(* PLC project station_cds.project, CODESYS CODESYS V3.5 SP22 Patch 1 *)
(* stored: creationDateTime 2026-11-25T17:27:32.1859428, modificationDateTime 2026-11-25T17:27:31.3827148 *)

FUNCTION_BLOCK FB_CurveEval
  VAR_INPUT
    Reset : BOOL;  (* clear all results, before a new pull *)
    Sample : BOOL;  (* X and F are a new sample *)
    Stroke : INT;  (* 1 pull, 2 return *)
    X : REAL;  (* mm, travel from touch *)
    F : REAL;  (* N *)
    Finish : BOOL;  (* return stroke finished: judge *)
    Mode : INT := 3;
    GateX : REAL := 3.0;  (* mm *)
    Gate2X : REAL := 10.0;  (* mm *)
    PeakXLo : REAL := 13.0;  (* mm *)
    PeakXHi : REAL := 26.0;  (* mm *)
    StepSpan : REAL := 2.0;  (* mm *)
    StopF : REAL := 30.0;  (* N *)
    G1Lo : REAL;  (* N, limits of FpG1 (mode 2) *)
    G1Hi : REAL;
    MeanLo : REAL;  (* N, limits of FMean (mode 3) *)
    MeanHi : REAL;
    HystLo : REAL;  (* N, limits of FHyst (mode 3) *)
    HystHi : REAL;
    RetFMin : REAL;  (* N, FrG1 must be above (mode 3) *)
    G2Lo : REAL;  (* N, limits of FpG2 *)
    G2Hi : REAL;
    PeakFLo : REAL;  (* N *)
    PeakFHi : REAL;
    PeakXMin : REAL;  (* mm, limits of XPeak *)
    PeakXMax : REAL;
    StepLo : REAL;  (* N *)
    StopXLo : REAL;  (* mm *)
    StopXHi : REAL;
    EnvX0 : REAL := 1.0;  (* mm, first envelope node *)
    EnvDx : REAL := 0.5;  (* mm, node spacing *)
    EnvN : INT := 55;  (* number of nodes, at most 64 *)
    EnvLo : ARRAY[0..63] OF REAL;  (* N *)
    EnvHi : ARRAY[0..63] OF REAL;  (* N *)
  END_VAR
  VAR_OUTPUT
    FpG1 : REAL;
    FrG1 : REAL;
    FMean : REAL;
    FHyst : REAL;
    FpG2 : REAL;
    FPeak : REAL;
    XPeak : REAL;
    FStep : REAL;
    XStop : REAL;
    EnvViol : INT;  (* envelope nodes outside the band *)
    EnvNodes : INT;  (* envelope nodes evaluated *)
    NSamples : INT;
    Done : BOOL;
    Ok : BOOL;
    NokCode : INT;
  END_VAR
  VAR
    sHavePrev : BOOL;
    sPrevX : REAL;
    sPrevF : REAL;
    sPrevStroke : INT;
    sGotG1 : BOOL;
    sGotG2 : BOOL;
    sGotR1 : BOOL;
    sGotPeak : BOOL;
    sGotStop : BOOL;
    sFMin : REAL;
    sFpG1 : REAL;
    sFrG1 : REAL;
    sFMean : REAL;
    sFHyst : REAL;
    sFpG2 : REAL;
    sFPeak : REAL;
    sXPeak : REAL;
    sFStep : REAL;
    sXStop : REAL;
    sEnvViol : INT;
    sEnvNodes : INT;
    sNSamples : INT;
    sDone : BOOL;
    sOk : BOOL;
    sNokCode : INT;
  END_VAR
  VAR_TEMP
    tI : INT;
    tNodeX : REAL;
    tFn : REAL;
    tCode : INT;
  END_VAR

                {region "Reset"}
        IF Reset THEN
            sFpG1 := 0.0;
            sFrG1 := 0.0;
            sFMean := 0.0;
            sFHyst := 0.0;
            sFpG2 := 0.0;
            sFPeak := 0.0;
            sXPeak := 0.0;
            sFStep := 0.0;
            sXStop := 0.0;
            sEnvViol := 0;
            sEnvNodes := 0;
            sNSamples := 0;
            sDone := FALSE;
            sOk := FALSE;
            sNokCode := 0;
            sHavePrev := FALSE;
            sGotG1 := FALSE;
            sGotG2 := FALSE;
            sGotR1 := FALSE;
            sGotPeak := FALSE;
            sGotStop := FALSE;
            sFMin := 0.0;
        END_IF;
    {endregion}

    {region "PullStroke"}
        IF NOT Reset AND Sample AND NOT sDone AND Stroke = 1 THEN
            IF sHavePrev AND sPrevStroke = 1 THEN
                // gates: force at a set travel, linear between the two samples around it
                IF NOT sGotG1 AND sPrevX < GateX AND X >= GateX THEN
                    sFpG1 := sPrevF + (F - sPrevF) * (GateX - sPrevX) / (X - sPrevX);
                    sGotG1 := TRUE;
                END_IF;
                IF NOT sGotG2 AND sPrevX < Gate2X AND X >= Gate2X THEN
                    sFpG2 := sPrevF + (F - sPrevF) * (Gate2X - sPrevX) / (X - sPrevX);
                    sGotG2 := TRUE;
                END_IF;
                // end stop: travel at a set force
                IF NOT sGotStop AND sPrevX > Gate2X AND sPrevF < StopF AND F >= StopF THEN
                    sXStop := sPrevX + (X - sPrevX) * (StopF - sPrevF) / (F - sPrevF);
                    sGotStop := TRUE;
                END_IF;
                // envelope: at most four nodes can lie between two samples
                FOR tI := 1 TO 4 DO
                    tNodeX := EnvX0 + EnvDx * INT_TO_REAL(sEnvNodes);
                    IF sEnvNodes < EnvN AND sPrevX < tNodeX AND X >= tNodeX THEN
                        tFn := sPrevF + (F - sPrevF) * (tNodeX - sPrevX) / (X - sPrevX);
                        IF tFn < EnvLo[sEnvNodes] OR tFn > EnvHi[sEnvNodes] THEN
                            sEnvViol := sEnvViol + 1;
                        END_IF;
                        sEnvNodes := sEnvNodes + 1;
                    END_IF;
                END_FOR;
            END_IF;
            // latch release: peak inside the window, then the drop after it
            IF X >= PeakXLo AND X <= PeakXHi AND (NOT sGotPeak OR F > sFPeak) THEN
                sFPeak := F;
                sXPeak := X;
                sFMin := F;
                sGotPeak := TRUE;
            ELSIF sGotPeak AND X <= sXPeak + StepSpan AND F < sFMin THEN
                sFMin := F;
            END_IF;
            IF sGotPeak THEN
                sFStep := sFPeak - sFMin;
            END_IF;
        END_IF;
    {endregion}

    {region "ReturnStroke"}
        IF NOT Reset AND Sample AND NOT sDone AND Stroke = 2 AND sHavePrev THEN
            IF NOT sGotR1 AND sPrevX > GateX AND X <= GateX THEN
                sFrG1 := sPrevF + (F - sPrevF) * (GateX - sPrevX) / (X - sPrevX);
                sGotR1 := TRUE;
            END_IF;
        END_IF;
    {endregion}

    {region "Bookkeeping"}
        IF NOT Reset AND Sample AND NOT sDone THEN
            sPrevX := X;
            sPrevF := F;
            sPrevStroke := Stroke;
            sHavePrev := TRUE;
            IF sNSamples < 32000 THEN
                sNSamples := sNSamples + 1;
            END_IF;
        END_IF;
    {endregion}

    {region "Verdict"}
        IF NOT Reset AND Finish AND NOT sDone THEN
            sFMean := (sFpG1 + sFrG1) * 0.5;
            sFHyst := sFpG1 - sFrG1;
            tCode := 0;
            CASE Mode OF
                1:  // peak force only
                    IF NOT sGotPeak THEN
                        tCode := 1;
                    ELSIF sFPeak < PeakFLo OR sFPeak > PeakFHi THEN
                        tCode := 6;
                    END_IF;
                2, 3:  // windows; mode 3 judges gate 1 with the return stroke
                    IF NOT (sGotG1 AND sGotG2 AND sGotPeak AND sGotStop) THEN
                        tCode := 1;
                    ELSIF Mode = 3 AND NOT sGotR1 THEN
                        tCode := 1;
                    ELSIF Mode = 2 AND (sFpG1 < G1Lo OR sFpG1 > G1Hi) THEN
                        tCode := 2;
                    ELSIF Mode = 3 AND (sFMean < MeanLo OR sFMean > MeanHi) THEN
                        tCode := 2;
                    ELSIF Mode = 3 AND (sFHyst < HystLo OR sFHyst > HystHi) THEN
                        tCode := 3;
                    ELSIF Mode = 3 AND sFrG1 < RetFMin THEN
                        tCode := 4;
                    ELSIF sFpG2 < G2Lo OR sFpG2 > G2Hi THEN
                        tCode := 5;
                    ELSIF sFPeak < PeakFLo OR sFPeak > PeakFHi THEN
                        tCode := 6;
                    ELSIF sXPeak < PeakXMin OR sXPeak > PeakXMax THEN
                        tCode := 7;
                    ELSIF sFStep < StepLo THEN
                        tCode := 8;
                    ELSIF sXStop < StopXLo OR sXStop > StopXHi THEN
                        tCode := 9;
                    END_IF;
                4:  // envelope: every node reached and inside
                    IF sEnvNodes < EnvN THEN
                        tCode := 1;
                    ELSIF sEnvViol > 0 THEN
                        tCode := 10;
                    END_IF;
                ELSE
                    tCode := 1;
            END_CASE;
            sNokCode := tCode;
            sOk := tCode = 0;
            sDone := TRUE;
        END_IF;
    {endregion}

    {region "Outputs"}
        // the working values live in static variables; the outputs are written here and nowhere else
        FpG1 := sFpG1;
        FrG1 := sFrG1;
        FMean := sFMean;
        FHyst := sFHyst;
        FpG2 := sFpG2;
        FPeak := sFPeak;
        XPeak := sXPeak;
        FStep := sFStep;
        XStop := sXStop;
        EnvViol := sEnvViol;
        EnvNodes := sEnvNodes;
        NSamples := sNSamples;
        Done := sDone;
        Ok := sOk;
        NokCode := sNokCode;
    {endregion}

          
END_FUNCTION_BLOCK
